{attribute 'qualified_only'}
VAR_GLOBAL
    // Bumped by every FB_ModeNodeSpy scan, so a test can check call order.
    nScanCounter : DINT;
END_VAR

(* stored: Version 1.1.0.1
   GVL GVL_Test: Id {3306825f-7f01-4b85-9db2-389af851c0d0} *)
